FUNCTION_BLOCK FB_Light IMPLEMENTS I_Light
VAR_INPUT
    stDeviceId : ST_DeviceId;
    iRelay     : I_Relay;
END_VAR

// FB_Light delegates relay operations through I_Relay.

PROPERTY DeviceId : ST_DeviceId
GET
DeviceId := stDeviceId;
END_GET
END_PROPERTY

PROPERTY IsOn : BOOL
GET
IsOn := iRelay.IsOn;
END_GET
END_PROPERTY

METHOD PUBLIC TurnOn
iRelay.TurnOn();
END_METHOD

METHOD PUBLIC TurnOff
iRelay.TurnOff();
END_METHOD

METHOD PUBLIC Toggle
iRelay.Toggle();
END_METHOD

METHOD PUBLIC SetBrightness
VAR_INPUT
    nBrightness : UINT;
END_VAR
// A relay-backed light supports only on/off switching.
// Zero switches it off; any non-zero level switches it on.
// A dimmer-backed light implementation can provide actual level control.
IF nBrightness = 0 THEN
    iRelay.TurnOff();
ELSE
    iRelay.TurnOn();
END_IF
END_METHOD

END_FUNCTION_BLOCK

(* stored: Version 1.1.0.1, ProductVersion 3.1.4026.20
   POU FB_Light: Id {B2B2B2B2-B2B2-42B2-82B2-B2B2B2B2B2B0}
   Property DeviceId: Id {B2B2B2B2-B2B2-42B2-82B2-B2B2B2B2B2B1}
   Get Get: Id {B2B2B2B2-B2B2-42B2-82B2-B2B2B2B2B2B2}
   Property IsOn: Id {B2B2B2B2-B2B2-42B2-82B2-B2B2B2B2B2B3}
   Get Get: Id {B2B2B2B2-B2B2-42B2-82B2-B2B2B2B2B2B4}
   Method TurnOn: Id {B2B2B2B2-B2B2-42B2-82B2-B2B2B2B2B2B5}
   Method TurnOff: Id {B2B2B2B2-B2B2-42B2-82B2-B2B2B2B2B2B6}
   Method Toggle: Id {B2B2B2B2-B2B2-42B2-82B2-B2B2B2B2B2B7}
   Method SetBrightness: Id {B2B2B2B2-B2B2-42B2-82B2-B2B2B2B2B2B8} *)
